(* IEC 61131-3 sources: brew/plant/generated/fleet/cs/openplc/cs-plc-utilities, 1 file *)

(* ---- located_vars.st ---- *)
(* Generated by plantgen from plant/plant.yaml and plant/sites.yaml (site cs). Do not edit. *)
(* Analog values are raw registers: engineering value = raw / 10^scaling. *)
(* RIO I/O is at %IX100.0 / %QX100.0 / %IW100 / %QW100 (v3 and v4 alike). *)
(* PLC memory: bits from %QX0.0 (coils), words from %MW0 (holding register qw_count and up, see modbus_slave.json). *)
VAR
  UTL_CHL_TT01_PV AT %IW100 : UINT; (* Glycol supply temperature, degF, x10 *)
  UTL_CHL_TT01_ALM_HIGH AT %QX0.0 : BOOL; (* Glycol supply temperature: high alarm (high) *)
  UTL_CHL_TT02_PV AT %IW101 : UINT; (* Glycol return temperature, degF, x10 *)
  UTL_CHL_JT01_PV AT %IW102 : UINT; (* Chiller electrical input, kW, x10 *)
  UTL_CHL_YS01_PV AT %IX100.0 : BOOL; (* Compressor stage 1 running *)
  UTL_CHL_YS02_PV AT %IX100.1 : BOOL; (* Compressor stage 2 running *)
  UTL_CHL_YA01_PV AT %IX100.2 : BOOL; (* Chiller compressor fault *)
  UTL_CHL_YA01_ALM_STATE AT %QX0.1 : BOOL; (* Chiller compressor fault: state alarm (high) *)
  UTL_CHL_HS01_CMD AT %QX100.0 : BOOL; (* Chiller enable *)
  UTL_CHL_TIC01_SP AT %QW100 : UINT; (* Chiller supply setpoint (written to the OEM controller), degF, x10 *)
  UTL_CHL_AT01_PV AT %IW103 : UINT; (* Refrigerant detector at the chiller (R-410A, 45 lb charge; ASHRAE 15), ppm, x1 *)
  UTL_CHL_AT01_ALM_HIGH AT %QX0.2 : BOOL; (* Refrigerant detector at the chiller (R-410A, 45 lb charge; ASHRAE 15): high alarm (high) *)
  UTL_CHL_TT01_SP AT %MW0 : UINT; (* Glycol supply setpoint (operator), degF, x10 *)
  UTL_GLY_LT01_PV AT %IW104 : UINT; (* Glycol reservoir level, %, x10 *)
  UTL_GLY_LT01_ALM_LOW AT %QX0.3 : BOOL; (* Glycol reservoir level: low alarm (medium) *)
  UTL_GLY_PT01_PV AT %IW105 : UINT; (* Glycol supply pressure, psig, x10 *)
  UTL_GLY_YS01_PV AT %IX100.3 : BOOL; (* Glycol pump running *)
  UTL_GLY_HS01_CMD AT %QX100.1 : BOOL; (* Glycol pump run command *)
  UTL_GLY_SC01_OUT AT %QW101 : UINT; (* Glycol pump VFD speed reference (pressure control), %, x10 *)
  UTL_GLY_PT01_SP AT %MW1 : UINT; (* Glycol supply pressure setpoint, psig, x10 *)
  UTL_STM_PT01_PV AT %IW106 : UINT; (* Steam header pressure, psig, x10 *)
  UTL_STM_PT01_ALM_LOW AT %QX0.4 : BOOL; (* Steam header pressure: low alarm (medium) *)
  UTL_STM_JT01_PV AT %IW107 : UINT; (* Boiler electrical input, kW, x10 *)
  UTL_STM_YS01_PV AT %IX100.4 : BOOL; (* Boiler firing *)
  UTL_STM_LSL01_PV AT %IX100.5 : BOOL; (* Boiler low-water cutoff tripped (hardwired) *)
  UTL_STM_LSL01_ALM_STATE AT %QX0.5 : BOOL; (* Boiler low-water cutoff tripped (hardwired): state alarm (high) *)
  UTL_STM_HS01_CMD AT %QX100.2 : BOOL; (* Boiler enable *)
  UTL_STM_PC01_SP AT %QW102 : UINT; (* Boiler pressure setpoint (12 psig; below the 15 psig safety valve), psig, x10 *)
  UTL_AIR_PT01_PV AT %IW108 : UINT; (* Compressed-air header pressure, psig, x10 *)
  UTL_AIR_PT01_ALM_LOW AT %QX0.6 : BOOL; (* Compressed-air header pressure: low alarm (medium) *)
  UTL_AIR_YS01_PV AT %IX100.6 : BOOL; (* Air compressor running *)
  UTL_AIR_YA01_PV AT %IX100.7 : BOOL; (* Air dryer fault *)
  UTL_AIR_HS01_CMD AT %QX100.3 : BOOL; (* Air compressor enable *)
  UTL_CO2_PT01_PV AT %IW109 : UINT; (* Bulk CO2 tank pressure, psig, x10 *)
  UTL_CO2_LT01_PV AT %IW110 : UINT; (* Bulk CO2 tank level, %, x10 *)
  UTL_CO2_LT01_ALM_LOW AT %QX0.7 : BOOL; (* Bulk CO2 tank level: low alarm (low) *)
  UTL_CO2_PT02_PV AT %IW111 : UINT; (* CO2 supply header pressure, psig, x10 *)
  UTL_CO2_PT02_ALM_LOW AT %QX1.0 : BOOL; (* CO2 supply header pressure: low alarm (medium) *)
  UTL_CO2_XV01_CMD AT %QX100.4 : BOOL; (* CO2 main supply valve (fail closed; its solenoid is wired through the shutoff relay) *)
  UTL_CO2_ZSO01_PV AT %IX101.0 : BOOL; (* CO2 main supply valve open (limit switch) *)
  UTL_CO2_XS01_CO2_OK AT %IX101.1 : BOOL; (* CO2 shutoff relay healthy (every area below 30,000 ppm, detection powered) *)
  UTL_CO2_XS02_SHUTOFF AT %QX1.1 : BOOL; (* CO2 supply shut off (tier 3 or loss of detection; latched until reset) *)
  UTL_CO2_XS02_ALM_STATE AT %QX1.2 : BOOL; (* CO2 supply shut off (tier 3 or loss of detection; latched until reset): state alarm (high) *)
  UTL_CO2_XC01_RESET AT %QX1.3 : BOOL; (* CO2 supply shutoff reset (operator; accepted once the relay has been healthy for 60 s) *)
  UTL_RO_FT01_PV AT %IW112 : UINT; (* RO permeate flow, gal/min, x10 *)
  UTL_RO_AT01_PV AT %IW113 : UINT; (* RO permeate conductivity, uS/cm, x1 *)
  UTL_RO_AT01_ALM_HIGH AT %QX1.4 : BOOL; (* RO permeate conductivity: high alarm (low) *)
  UTL_RO_YS01_PV AT %IX101.2 : BOOL; (* RO skid running *)
  UTL_RO_HS01_CMD AT %QX100.5 : BOOL; (* RO skid run command *)
  UTL_WWN_LT01_PV AT %IW114 : UINT; (* Neutralization tank level, %, x10 *)
  UTL_WWN_LT01_ALM_HIGH AT %QX1.5 : BOOL; (* Neutralization tank level: high alarm (medium) *)
  UTL_WWN_AT01_PV AT %IW115 : UINT; (* Neutralization tank pH, pH, x100 *)
  UTL_WWN_AT01_ALM_HIGH AT %QX1.6 : BOOL; (* Neutralization tank pH: high alarm (low) *)
  UTL_WWN_AT01_ALM_LOW AT %QX1.7 : BOOL; (* Neutralization tank pH: low alarm (low) *)
  UTL_WWN_LSH01_PV AT %IX101.3 : BOOL; (* Neutralization tank high-level switch *)
  UTL_WWN_XV01_CMD AT %QX100.6 : BOOL; (* Caustic dosing pump *)
  UTL_WWN_XV02_CMD AT %QX100.7 : BOOL; (* Acid dosing pump *)
  UTL_WWN_XV03_CMD AT %QX101.0 : BOOL; (* Discharge valve to the sewer (permitted at pH 6.0-9.0) *)
  UTL_WWN_XS01_INHIBIT AT %QX2.0 : BOOL; (* Discharge inhibited (pH outside 6.0-9.0) *)
  UTL_WWN_XS01_ALM_STATE AT %QX2.1 : BOOL; (* Discharge inhibited (pH outside 6.0-9.0): state alarm (medium) *)
  UTL_CIP_TT01_PV AT %IW116 : UINT; (* CIP supply temperature, degF, x10 *)
  UTL_CIP_TT01_ALM_DEVIATION AT %QX2.2 : BOOL; (* CIP supply temperature: deviation alarm (low) *)
  UTL_CIP_AT01_PV AT %IW117 : UINT; (* CIP return conductivity, mS/cm, x100 *)
  UTL_CIP_FT01_PV AT %IW118 : UINT; (* CIP return flow, gal/min, x10 *)
  UTL_CIP_LT01_PV AT %IW119 : UINT; (* Caustic tank level, %, x10 *)
  UTL_CIP_LT02_PV AT %IW120 : UINT; (* Acid/sanitizer tank level, %, x10 *)
  UTL_CIP_FS01_PV AT %IX101.4 : BOOL; (* CIP return flow proven (flow switch) *)
  UTL_CIP_HS01_CMD AT %QX101.1 : BOOL; (* CIP supply pump run command *)
  UTL_CIP_HS02_CMD AT %QX101.2 : BOOL; (* CIP return pump run command *)
  UTL_CIP_XV01_CMD AT %QX101.3 : BOOL; (* Caustic dosing *)
  UTL_CIP_XV02_CMD AT %QX101.4 : BOOL; (* Acid/sanitizer dosing *)
  UTL_CIP_TV01_OUT AT %QW103 : UINT; (* CIP heater steam valve position, %, x10 *)
  UTL_CIP_ZS01_PV AT %IX101.5 : BOOL; (* Swing panel on the brewhouse circuit *)
  UTL_CIP_ZS02_PV AT %IX101.6 : BOOL; (* Swing panel on FV-101 *)
  UTL_CIP_ZS03_PV AT %IX101.7 : BOOL; (* Swing panel on FV-102 *)
  UTL_CIP_ZS04_PV AT %IX102.0 : BOOL; (* Swing panel on FV-103 *)
  UTL_CIP_ZS05_PV AT %IX102.1 : BOOL; (* Swing panel on FV-104 *)
  UTL_CIP_ZS06_PV AT %IX102.2 : BOOL; (* Swing panel on BBT-201 *)
  UTL_CIP_ZS07_PV AT %IX102.3 : BOOL; (* Swing panel on BBT-202 *)
  UTL_CIP_TT01_SP AT %MW2 : UINT; (* CIP supply temperature setpoint, degF, x10 *)
  UTL_CIP_XC01_CIRCUIT AT %MW3 : UINT; (* CIP circuit selected (1 to 7; 0 none), None, x1 *)
  UTL_CIP_XC01_CMD AT %MW4 : UINT; (* CIP sequence command (1 start, 2 hold, 3 abort), None, x1 *)
  UTL_CIP_XS01_STEP AT %MW5 : UINT; (* CIP sequence step, None, x1 *)
  UTL_CIP_XS02_ROUTE_OK AT %QX2.3 : BOOL; (* CIP route verified (the swing panel is on the circuit and the cellar permits it) *)
  UTL_CIP_XS03_PV AT %IX120.0 : BOOL; (* Cellar transfer in progress (peer read from cs-plc-cellar) *)
  UTL_CIP_XS04_PV AT %IX120.1 : BOOL; (* Cellar circuits permit CIP (peer read from cs-plc-cellar) *)
  UTL_CIP_XS05_PV AT %IX120.2 : BOOL; (* FV-101 not in entry (peer read from cs-plc-cellar) *)
  UTL_CIP_XS06_PV AT %IX120.3 : BOOL; (* FV-102 not in entry (peer read from cs-plc-cellar) *)
  UTL_CIP_XS07_PV AT %IX120.4 : BOOL; (* FV-103 not in entry (peer read from cs-plc-cellar) *)
  UTL_CIP_XS08_PV AT %IX120.5 : BOOL; (* FV-104 not in entry (peer read from cs-plc-cellar) *)
  UTL_CIP_XS09_PV AT %IX120.6 : BOOL; (* BBT-201 not in entry (peer read from cs-plc-cellar) *)
  UTL_CIP_XS10_PV AT %IX120.7 : BOOL; (* BBT-202 not in entry (peer read from cs-plc-cellar) *)
  UTL_CIP_XA01_PV AT %QX2.4 : BOOL; (* CIP held: return flow lost (the pumps stay off until Hold and Resume, or Abort) *)
  UTL_CIP_XA01_ALM_STATE AT %QX2.5 : BOOL; (* CIP held: return flow lost (the pumps stay off until Hold and Resume, or Abort): state alarm (medium) *)
END_VAR
